FUNCTION_BLOCK TankModel IMPLEMENTS I_LevelSensor, I_Cyclic
VAR
    _Inflow       : I_FillValve;
    _Outflow      : I_FillValve;
    _Clock        : I_Clock;
    _FillRate     : REAL;              // percent per second, inflow valve open
    _DrainRate    : REAL;              // percent per second, outflow valve open
    _Level        : REAL;
    _LastNow      : LTIME;
    _IsStarted    : BOOL;
    _IsConfigured : BOOL;
END_VAR
(*
    TankModel

    A simulated tank: the level rises while the inflow valve is open and
    falls while the outflow valve is open. Reads both through
    I_FillValve, so it works with simulated and real valves alike.
*)

METHOD FB_init : BOOL
VAR_INPUT
    bInitRetains : BOOL;
    bInCopyCode  : BOOL;
    Inflow       : I_FillValve;
    Outflow      : I_FillValve;
    Clock        : I_Clock;
    FillRate     : REAL;
    DrainRate    : REAL;
    StartLevel   : REAL;
END_VAR
_Inflow := Inflow;
_Outflow := Outflow;
_Clock := Clock;
_FillRate := FillRate;
_DrainRate := DrainRate;
_Level := StartLevel;
_IsConfigured := Inflow <> 0 AND Outflow <> 0 AND Clock <> 0;
END_METHOD

METHOD PUBLIC CyclicLogic
VAR
    Now     : LTIME;
    Seconds : REAL;
END_VAR
IF NOT _IsConfigured THEN
    RETURN;
END_IF
Now := _Clock.Now;
IF NOT _IsStarted THEN
    _IsStarted := TRUE;
    _LastNow := Now;
    RETURN;
END_IF
Seconds := LREAL_TO_REAL(LTIME_TO_LREAL(Now - _LastNow) / 1.0E9);   // LTIME counts nanoseconds
_LastNow := Now;
IF _Inflow.IsOpen THEN
    _Level := _Level + _FillRate * Seconds;
END_IF
IF _Outflow.IsOpen THEN
    _Level := _Level - _DrainRate * Seconds;
END_IF
_Level := LIMIT(0.0, _Level, 100.0);
END_METHOD

PROPERTY PUBLIC Level : REAL
GET
Level := _Level;
END_GET
END_PROPERTY

PROPERTY PUBLIC IsValid : BOOL
GET
IsValid := _IsConfigured;
END_GET
END_PROPERTY

END_FUNCTION_BLOCK

(* stored: Version 1.1.0.1, ProductVersion 3.1.4026.0
   POU TankModel: Id {7e8c216c-b31a-4907-b57b-4834cc757592}, SpecialFunc None
   Folder I_LevelSensor: Id {e48ccde3-8e33-40cf-b794-3ff9a0b9226a}
   Folder I_Cyclic: Id {274ca545-2b3a-41d7-bd13-1d203c19f46f}
   Method FB_init: Id {e5a14c5e-8902-4b9d-a9a3-be269beee06f}
   Method CyclicLogic: Id {2209cb73-3c89-40af-8de4-a1f136a4f553}
   Property Level: Id {916f4c91-a9f9-486c-b73b-270876f42d1f}
   Get Get: Id {35e616ea-8034-4aea-8855-2ffe9047b042}
   Property IsValid: Id {44624941-7c11-482a-8e63-0b5e383fdeb1}
   Get Get: Id {626b1e44-dcb7-45ae-aea6-ffa8ab07c505} *)
